Fanuc KAREL source: KT00707.KL

PROGRAM KT00707
%NOLOCKGROUP
VAR
  I1: INTEGER
  I2: INTEGER
  OUT: INTEGER
BEGIN
  I1 = 2
  I2 = 3
  I1 = 2
  I2 = 3
  OUT = ARRAY_LEN(I1)
END KT00707
